(* IEC 61131-3 sources: plc-process-lib/tests/POUs/Helpers/FB_TestSink, 4 files *)

(* ---- FB_TestSink.decl.st ---- *)
// Назначение: тестовый приёмник событий тревог (I_AlarmSink): кольцо на 32 события.
//             Подставляется в GVL_Lib.itfAlarmSink только в тестах, которым нужны события;
//             тест возвращает GVL_Lib.itfAlarmSink := 0 до coUnit.TEST_FINISHED().
// Автор:      kr0nsch
// Версия:     0.1.0
// Документ:   docs/TESTING.md, раздел «Вспомогательные ФБ»
FUNCTION_BLOCK FB_TestSink IMPLEMENTS I_AlarmSink
VAR CONSTANT
    EVENTS_MAX : UINT := 32;                   // ёмкость кольца
END_VAR
VAR
    astEvent : ARRAY[0..EVENTS_MAX - 1] OF ST_AlarmEvent;  // кольцо событий
    uiNext   : UINT;                           // индекс следующей записи
    uiCount  : UINT;                           // событий с последнего Clear (не больше UINT_MAX)
END_VAR

(* ---- GetEvent.method.decl.st ---- *)
// Событие, записанное uiBack событий назад (0 — последнее); нет такого — пустое событие
METHOD PUBLIC GetEvent : ST_AlarmEvent
VAR_INPUT
    uiBack : UINT;             // сколько событий назад
END_VAR
VAR
    stNone : ST_AlarmEvent;    // пустое событие
END_VAR

(* ---- GetEvent.method.impl.st ---- *)
IF uiBack < MIN(uiCount, EVENTS_MAX) THEN
    GetEvent := astEvent[(uiNext + EVENTS_MAX - 1 - uiBack) MOD EVENTS_MAX];
ELSE
    GetEvent := stNone;
END_IF

(* ---- OnAlarmEvent.method.decl.st ---- *)
// Записать событие в кольцо (самое старое затирается); приёмник не переполняется — TRUE
METHOD PUBLIC OnAlarmEvent : BOOL
VAR_IN_OUT CONSTANT
    stEvent : ST_AlarmEvent;   // событие
END_VAR
